Fanuc KAREL source: kt00343.KL

-- PROVISIONAL review KL for V1013-1; original PC SHA256 8168a37a1c84f3df904550553125e70268de4978b0cd3114442241ec26dc3df9
-- Incomplete behavior may be omitted. Consult companion uncertainty JSON. Do not deploy.
PROGRAM KT00343
%NOLOCKGROUP
VAR
  I2 : INTEGER
  OUT : BOOLEAN
-- UNRESOLVED_DECL H1 type=002017
BEGIN
  -- UNRESOLVED_PC offsets 5-19; opcodes 2E,22,9D,33,B4
  -- UNRESOLVED_PC offsets 24-35; opcodes 2E,23
  -- UNRESOLVED_PC offsets 40-62; opcodes 22,9D,33,B3,21,59,23
  -- UNRESOLVED_PC offsets 67-71; opcodes 7F
END KT00343
